(* IEC 61131-3 sources: plc-workbench/examples/motor, 2 files *)

(* ---- alternative.st ---- *)
FUNCTION_BLOCK MotorControl
VAR_INPUT
    StartBtn : BOOL;
    StopBtn : BOOL;
    EStop : BOOL;
END_VAR
VAR_OUTPUT
    Motor : BOOL := FALSE;
END_VAR
Motor := (Motor OR StartBtn) AND NOT StopBtn AND NOT EStop;
END_FUNCTION_BLOCK

(* ---- correct.st ---- *)
FUNCTION_BLOCK MotorControl
VAR_INPUT
    StartBtn : BOOL;
    StopBtn : BOOL;
    EStop : BOOL;
END_VAR
VAR_OUTPUT
    Motor : BOOL := FALSE;
END_VAR
IF StopBtn OR EStop THEN
    Motor := FALSE;
ELSIF StartBtn THEN
    Motor := TRUE;
END_IF;
END_FUNCTION_BLOCK
